// TIA Portal V21 export
// export: Created 2026-11-22T04:06:10.5650757Z, ExportSetting WithDefaults, DisplayName Totally Integrated Automation Portal, DisplayVersion V21 Update 3, DisplayName STEP 7 Professional, DisplayVersion V21 Update 3, DisplayName STEP 7 Safety, DisplayVersion V21, DisplayName Tech WebApplication, DisplayVersion V21, DisplayName WinCC Basic/Comfort/Advanced, DisplayVersion V21 Update 3, DisplayName WinCC Unified, DisplayVersion V21 Update 3
ScreenTemplate "T_C05"  1280x800
  ScreenLayer "Layer_0"
    Rectangle "T_Header" at 0,0 size 1280x34
    TextField "T_Title" at 8,6 size 300x22  Text="Template T_C05 (header)"
    DateTimeField "T_Clock" at 1090,4 size 180x26  Mode=Output
